Fanuc KAREL source: kt00567.KL

-- PROVISIONAL review KL for V1013-1; original PC SHA256 e03df45c199e0e37e2bfcf72bbef2f9e0064e12c007617a87b26523f9f4caf05
-- Incomplete behavior may be omitted. Consult companion uncertainty JSON. Do not deploy.
PROGRAM KT00567
%NOLOCKGROUP
VAR
  R2 : REAL
-- UNRESOLVED_DECL V1 type=000013
-- UNRESOLVED_DECL OUT type=000013
BEGIN
  -- UNRESOLVED_PC offsets 5-20; opcodes 2E,22,32,35
  -- UNRESOLVED_PC offsets 25-36; opcodes 2E,23
  -- UNRESOLVED_PC offsets 41-63; opcodes 49,21,8A,4A
  -- UNRESOLVED_PC offsets 68-72; opcodes 7F
END KT00567
